(* PLC project coil_on_input, ESBMC probe 1.0 *)
(* stored: creationDateTime 2026-10-07T00:00:00 *)

PROGRAM coil_on_input
  VAR_INPUT
    x : BOOL;
    go : BOOL;
  END_VAR
  VAR_OUTPUT
    q : BOOL;
  END_VAR

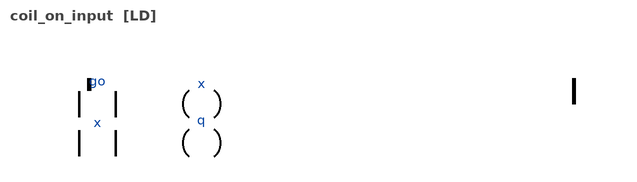
(* LD diagram, written out as Structured Text *)
x := go;
q := x;
END_PROGRAM

CONFIGURATION Config0
  RESOURCE Res0 ON PLC
    TASK tcyclic(INTERVAL := T#10ms, PRIORITY := 0);
    PROGRAM inst0 WITH tcyclic : coil_on_input;
  END_RESOURCE
END_CONFIGURATION
